(* IEC 61131-3 sources: 2026_Projet_YGO_ExcavatriceDragage/CODE/G_CYCLE (part 3) *)

    E_AutoCycleStep.AX15A_DUMP_ARRIVE:
        CycleStep := E_AutoCycleStep.AX15A_DUMP_ARRIVE;
        CycleStateStr := 'AX15a - Arrivee tremie : treuils arretes, attente ouverture';
        Lifecycle.Busy := TRUE;
        Lifecycle.Done := FALSE;
        ExpectedAxis := E_OperatorAxis.JOYSTICK_Y;
        ExpectedDirection := -1;
        WaitingForOperator := TRUE;
        WaitingForProcess := FALSE;
        OperatorActionId := 16#040B;
        OperatorAction := 'AX15a - Relacher le joystick avant ouverture.';

        // Config treuil UNIQUE : arret des deux treuils (aucune descente couplee ici).
        WinchM1Cmd.RunRequest := FALSE; WinchM1Cmd.ReqAscent := FALSE; WinchM1Cmd.ReqDescend := FALSE; WinchM1Cmd.StepTgt := 0;
        WinchM2Cmd.RunRequest := FALSE; WinchM2Cmd.ReqAscent := FALSE; WinchM2Cmd.ReqDescend := FALSE; WinchM2Cmd.StepTgt := 0;
        TranslationCmd.ReqStart := FALSE;
        TranslationCmd.PositionTgt := 0;

        IF PvDumpLatched THEN
            BucketCmd.ReqOpen := DeadmanArmed AND JoystickPush;
        END_IF;

        IF PvDumpLatched AND Benne_Done AND Benne_IsOpen THEN
            BucketCmd.ReqOpen := FALSE;
            State := E_AutoCycleStep.AX18_DONE_SYNC;
        ELSIF (CfgPauseBeforeDump_S > 0.0) AND NOT PauseBeforeDumpTimer.Q THEN
            WaitingForOperator := FALSE;
            WaitingForProcess := TRUE;
            OperatorAction := 'AX15a - Stabilisation chariot avant ouverture benne.';
            IF NOT JoystickDeflected THEN
                SeenNeutralAfterArrival := TRUE;
            END_IF;
        ELSIF SeenNeutralAfterArrival OR PvDumpLatched THEN
            WaitingForOperator := NOT (DeadmanArmed AND JoystickPush);
            WaitingForProcess := DeadmanArmed AND JoystickPush;
            OperatorAction := 'AX15a - Pousser vers le bas pour ouvrir et vider.';
            IF DeadmanArmed AND JoystickPush THEN
                State := E_AutoCycleStep.AX15B_DUMP_OPEN;
            END_IF;
        ELSIF NOT JoystickDeflected THEN
            SeenNeutralAfterArrival := TRUE;
            OperatorAction := 'AX15a - Pousser vers le bas pour ouvrir et vider.';
        END_IF;

    E_AutoCycleStep.AX15B_DUMP_OPEN:
        CycleStep := E_AutoCycleStep.AX15B_DUMP_OPEN;
        CycleStateStr := 'AX15b - Vidage : ouverture benne, treuils arretes';
        Lifecycle.Busy := TRUE;
        Lifecycle.Done := FALSE;
        ExpectedAxis := E_OperatorAxis.JOYSTICK_Y;
        ExpectedDirection := -1;
        WaitingForOperator := NOT (DeadmanArmed AND JoystickPush);
        WaitingForProcess := DeadmanArmed AND JoystickPush;
        OperatorActionId := 16#040B;
        OperatorAction := 'AX15b - Pousser : vidage. Tirer : fermer et remonter.';

        // Config treuil UNIQUE : etape benne seule, les deux treuils neutralises
        // (plus de descente couplee M1+M2 simultanee a l'ouverture benne -> plus
        // d'ecart M1/M2 volontaire ni de faux SafeStop concordance contacteurs).
        WinchM1Cmd.RunRequest := FALSE; WinchM1Cmd.ReqAscent := FALSE; WinchM1Cmd.ReqDescend := FALSE; WinchM1Cmd.StepTgt := 0;
        WinchM2Cmd.RunRequest := FALSE; WinchM2Cmd.ReqAscent := FALSE; WinchM2Cmd.ReqDescend := FALSE; WinchM2Cmd.StepTgt := 0;
        TranslationCmd.ReqStart := FALSE;
        TranslationCmd.PositionTgt := 0;

        BucketCmd.ReqOpen := DeadmanArmed AND JoystickPush;

        // Vidage benne en AX15B
        IF RepositionRequest THEN
            State := E_AutoCycleStep.AX15C_DUMP_REPOSITION;
        ELSIF DeadmanArmed AND JoystickPush AND Benne_Done AND Benne_IsOpen THEN
            BucketCmd.ReqOpen := FALSE;
            State := E_AutoCycleStep.AX18_DONE_SYNC;
        END_IF;

    E_AutoCycleStep.AX15C_DUMP_REPOSITION:
        CycleStep := E_AutoCycleStep.AX15C_DUMP_REPOSITION;
        CycleStateStr := 'AX15c - Repositionnement couple M1+M2 (aide vidange tremie)';
        Lifecycle.Busy := TRUE;
        Lifecycle.Done := FALSE;
        ExpectedAxis := E_OperatorAxis.JOYSTICK_Y;
        ExpectedDirection := -1;
        WaitingForOperator := NOT JoystickDeflected;
        WaitingForProcess := JoystickDeflected;
        OperatorActionId := 16#040C;
        OperatorAction := 'AX15c - Descente couplee M1+M2 ; relacher l option pour reprendre le vidage.';

        // Descente couplee M1+M2, palier lent, sous homme-mort. Commandes SYMETRIQUES
        // (meme sens, meme palier) -> FB_SyncDeviation actif, pas d'ecart volontaire.
        WinchM1Cmd.ReqAscent := FALSE; WinchM1Cmd.ReqDescend := TRUE;
        WinchM1Cmd.RunRequest := CycleMotionPermit;
        WinchM1Cmd.StepTgt := CST_StepSlow;
        WinchM2Cmd.ReqAscent := FALSE; WinchM2Cmd.ReqDescend := TRUE;
        WinchM2Cmd.RunRequest := CycleMotionPermit;
        WinchM2Cmd.StepTgt := CST_StepSlow;
        TranslationCmd.ReqStart := FALSE;
        TranslationCmd.PositionTgt := 0;

        // La benne reste ouverte pendant le repositionnement (on finit l'ouverture si besoin).
        BucketCmd.ReqOpen := CycleMotionPermit AND NOT Benne_IsOpen;

        // Retour a AX15B des que l'operateur relache l'option de repositionnement.
        IF NOT RepositionRequest THEN
            WinchM1Cmd.RunRequest := FALSE;
            WinchM2Cmd.RunRequest := FALSE;
            State := E_AutoCycleStep.AX15B_DUMP_OPEN;
        END_IF;

    E_AutoCycleStep.AX18_DONE_SYNC:
        CycleStep := E_AutoCycleStep.AX18_DONE_SYNC;
        CycleStateStr := 'AX18 - Passe terminee : aller en P1 pour recommencer';
        WinchM1Cmd.RunRequest := FALSE;
        WinchM2Cmd.RunRequest := FALSE;
        TranslationCmd.ReqStart := FALSE;
        Lifecycle.Done := TRUE;
        Lifecycle.Busy := FALSE;
        ExpectedAxis := E_OperatorAxis.JOYSTICK_X;
        ExpectedDirection := 1;
        WaitingForOperator := NOT (DeadmanArmed AND JoystickRight);
        WaitingForProcess := DeadmanArmed AND JoystickRight;
        OperatorActionId := 16#040D;
        OperatorAction := 'AX18 - Cycle termine. Aller en P1 (joystick a droite).';

        // Compteur de prélèvements (RETAIN) + durée du cycle — F2: cadré par front (1 seul par cycle)
        IF NOT SampleCountDone THEN
            SampleCount := SampleCount + 1;            // JOURNALIER (RAZ IHM/mode auto possible)
            SampleCountTotal := SampleCountTotal + 1;  // TOTALISATEUR : SEULE ecriture de toute l'application (gate G508)
            LastCycleDuration_Min := CurrentCycleElapsed_Min;  // fige la duree du cycle qui vient de s'achever
            LastCycleDuration_S   := CurrentCycleElapsed_S;
            SampleCountDone := TRUE;
        END_IF;

        // Rebouclage DIRECT sur AX2_TRANSLATE_P1 (GEL Q14) : la machine est deja
        // referencee, la passe suivante enchaine sur la translation P1 (pas de retour AX0).
        // Relance sur StartCycle OU FRONT joystick (geste franc) - pas sur simple maintien,
        // pour que AX18 (Lifecycle.Done + msg) soit reellement observable / tracable.
        IF StartEdge.Q OR (DeadmanArmed AND JoystickRight) THEN
            SampleCountDone := FALSE;
            Lifecycle.Done := FALSE;
            State := E_AutoCycleStep.AX2_TRANSLATE_P1;
        END_IF;

    E_AutoCycleStep.AX_STAB:
        CycleStep := E_AutoCycleStep.AX_STAB;
        CycleStateStr := 'STABILISATION - defaut cycle';
        WinchM1Cmd.RunRequest := FALSE; WinchM1Cmd.ReqAscent := FALSE; WinchM1Cmd.ReqDescend := FALSE;
        WinchM2Cmd.RunRequest := FALSE; WinchM2Cmd.ReqAscent := FALSE; WinchM2Cmd.ReqDescend := FALSE;
        TranslationCmd.ReqStart := FALSE;
        BucketCmd.ReqOpen := FALSE;
        BucketCmd.ReqClose := FALSE;
        BucketCmd.ReqKoboldMeasureEnable := FALSE;   // Coupure contacteur Kobold au repli defaut (0 ordre residuel)
        Lifecycle.Busy := FALSE;
        Lifecycle.Done := FALSE;
        ExpectedAxis := E_OperatorAxis.BUTTON;
        ExpectedDirection := 0;
        WaitingForOperator := TRUE;
        WaitingForProcess := FALSE;
        OperatorActionId := 16#0480;
        IF ResumeAfterFaultAvailable THEN
            OperatorAction := 'AX_STAB : cause disparue - Reprendre ou Abandonner.';
        ELSIF Translation_PosMaintenance AND NOT Translation_PosP1 THEN
            // Reprise boot : Maintenance active + P1 retombe = chariot déjà au-delà
            // de P1. Ne jamais proposer de continuer à droite vers Maintenance.
            // Le retour gauche traverse P1 ; le front P1 réarme AtP1 et la branche
            // précédente termine AX2 normalement.
            ExpectedDirection := 1;
            WaitingForOperator := NOT JoystickDeflected;
            WaitingForProcess := JoystickDeflected;
            OperatorActionId := 16#0402;
            OperatorAction := 'AX2 - M3 au-dela de P1 : pousser vers tremie (gauche) jusqu a P1.';
            TranslationCmd.PositionTgt := 1;      // sens retour vers Trémie
            TranslationCmd.ReqStart := TranslationTremiePermit;
        ELSE
            OperatorAction := 'AX_STAB : lever la cause puis Reprendre/Abandonner.';
        END_IF;

END_CASE;
END_IF;
{endregion}

{region "§4 Repli homme mort & Syntheses"}
// 🛑 Relâchement du manche (retour au centre) OU de l'homme-mort : neutralisation
// des demandes actives. Gate continu : aucune commande d'actionneur ne survit à la
// perte du permis opérateur (manche défléchi ET homme-mort armé).
IF Lifecycle.Busy AND NOT CycleMotionPermit THEN
    WinchM1Cmd.RunRequest := FALSE;
    WinchM2Cmd.RunRequest := FALSE;
    TranslationCmd.ReqStart := FALSE;
    BucketCmd.ReqOpen := FALSE;
    BucketCmd.ReqClose := FALSE;
    BucketCmd.ReqKoboldMeasureEnable := FALSE;
END_IF;

RequestActive := WinchM1Cmd.RunRequest OR WinchM2Cmd.RunRequest OR TranslationCmd.ReqStart OR BucketCmd.ReqOpen OR BucketCmd.ReqClose OR BucketCmd.ReqHoldAscentP1AfterClose OR BucketCmd.ReqKoboldMeasureEnable; // Somme logique complete des demandes (contacteur Kobold inclus)
{endregion}

END_FUNCTION_BLOCK
